TYPE ST_MenteeMotorV32OsSample :
STRUCT
    // Generic oversample slot (flex-PDO 0x6001). w0/w1/w2 are RAW 32-bit words for
    // the fixed lanes:  w0=theta(F)  w1=d_theta(F)  w2=iq(F)
    sample_idx  : UDINT;    // sN_sample_idx — device oversample index
    w0          : UDINT;    // sN_w0 — raw word (float bits)
    w1          : UDINT;    // sN_w1
    w2          : UDINT;    // sN_w2
    // Extended lanes 3..9 — ELF-picked debug variables on the slot-2 debug
    // pipe. Filled by FB_Slot2PipeHandler from the SAME
    // capture index k as w0..w2 (the FW samples every bound lane on one
    // shared prescaler tick), so one aSamples[k] is one synchronized instant
    // stamped by sample_idx. Stay 0 when no debug var is bound to that lane.
    w3          : UDINT;
    w4          : UDINT;
    w5          : UDINT;
    w6          : UDINT;
    w7          : UDINT;
    w8          : UDINT;
    w9          : UDINT;
END_STRUCT
END_TYPE

(* stored: Version 1.1.0.1, ProductVersion 3.1.4026.18
   DUT ST_MenteeMotorV32OsSample: Id {8d32101a-96bd-4154-848c-aeb8105ad132} *)
